// TIA Portal V21 export
// export: Created 2026-10-12T12:46:16.8935172Z, ExportSetting WithDefaults, DisplayName Totally Integrated Automation Portal, DisplayVersion V21, DisplayName STEP 7 Professional, DisplayVersion V21, DisplayName STEP 7 Safety, DisplayVersion V21, DisplayName Tech WebApplication, DisplayVersion V21, DisplayName WinCC Basic/Comfort/Advanced, DisplayVersion V21, DisplayName WinCC Unified, DisplayVersion V21
TagTable "Default tag table"
  Tag_ScreenNumber : UInt  (1 s)
  AUTO MODE SELECTED : Bool  (HMI_Connection_1, 1 s)
  DB_ALARMS_FAULT POP : Bool  (HMI_Connection_1, 1 s)
  DB_ALARMS_WARNING POP : Bool  (HMI_Connection_1, 1 s)
  DB_HMI_FAULT RESET PB : Bool  (HMI_Connection_1, 1 s)
  DB_HMI_MOTOR JOG FWD PB : Bool  (HMI_Connection_1, 1 s)
  DB_HMI_MOTOR JOG REV PB : Bool  (HMI_Connection_1, 1 s)
  DB_AUTO_AUTO STATUS : Int  (HMI_Connection_1, 1 s)
  DB_HMI_STOP TIME : DInt  (HMI_Connection_1, 1 s)
  DB_HMI_CAMERA DONE : Bool  (HMI_Connection_1, 1 s)
